(*
SPDX-FileCopyrightText: c 2026 Oleksandr Tiutyk <trofimich@gmail.com>
SPDX-License-Identifier: MIT
License: https://opensource.org/license/mit
*)

(*!
<summary>Checks that a long aggregate diagnostic is terminated and ends in an ellipsis.</summary>
<description>
Uses one task and stays at a stable address while assertions are bound to this instance.
</description>
*)

{attribute 'no_assign'}
{attribute 'no_explicit_call' := 'do not call this function block directly'}
FUNCTION_BLOCK AggregateExceptionBoundedMessageTest EXTENDS TOF_Testing.SingleCycleTest
VAR_STAT
	{attribute 'hide'}
	_ClassName : STRING := __POUNAME();
END_VAR
VAR
	_Aggregate : TOF_Core.AggregateException;
END_VAR

(*!
<summary>Checks that a long aggregate diagnostic is terminated and ends in an ellipsis.</summary>
<description>
Three entries share one task-managed cause. Each payload fills half the diagnostic buffer so the
combined message exceeds its capacity. The persistent reference array is released in AfterTest.
</description>
*)
METHOD PROTECTED ExecuteTest
VAR
	exceptionCode : __SYSTEM.ExceptionCode;
	caught : TOF_Core.IException;
	cause : TOF_Core.IStandardException;
	payload : TOF_Core.ERROR_MESSAGE;
	message : TOF_Core.ERROR_MESSAGE;
	payloadUnits : POINTER TO WORD;
	messageUnits : POINTER TO WORD;
	i : UDINT;
END_VAR
VAR CONSTANT
	MESSAGE_CAPACITY : UDINT := TOF_Core.Parameters.ERROR_MESSAGE_WIDE_CHAR_SIZE;
END_VAR
// Make an ASCII payload whose length scales with the documented diagnostic capacity.
payloadUnits := ADR(payload);

FOR i := 0 TO MESSAGE_CAPACITY / 2 - 1 DO
	payloadUnits[i] := WORD#16#0058; // Uppercase X makes the retained prefix distinguishable from the ellipsis.
END_FOR

payloadUnits[MESSAGE_CAPACITY / 2] := TO_WORD(TOF_Core.UnsignedInt16.MIN_VALUE);

// Obtain one dynamic cause so repeated entries exercise permitted sharing.
__TRY
	TOF_Core.Exceptions.ThrowStandard(
		sourceNamespaceName := NamespaceName,
		sourceClassName := ClassName,
		sourcePOUName := __POUNAME(),
		sourcePosition := __POSITION(),
		message := payload
	);
__CATCH(exceptionCode)
	caught := TOF_Core.ExceptionManager.GetLastException(
		exceptionCode := exceptionCode,
		catchPointNamespaceName := NamespaceName,
		catchPointPOUName := __POUNAME(),
		catchPointPosition := __POSITION()
	);
__ENDTRY

IF NOT __QUERYINTERFACE(caught, cause) THEN
	RecordFailure(message := "A task-owned payload is required for the aggregate length check");
	RETURN;
END_IF

_Aggregate.AddInnerException(innerException := cause);
_Aggregate.AddInnerException(innerException := cause);
_Aggregate.AddInnerException(innerException := cause);
message := _Aggregate.GetMessage();

messageUnits := ADR(message);

IF messageUnits[MESSAGE_CAPACITY] <> TO_WORD(TOF_Core.UnsignedInt16.MIN_VALUE) THEN
	RecordFailure(message := "The last storage unit must terminate the aggregate diagnostic");
	RETURN;
END_IF

Assert.ThatUDInt(
	actual := TOF_Core.WideStrings.GetLength(value := message),
	message := "The bounded aggregate message must fill the available character capacity"
).ToBe(expected := MESSAGE_CAPACITY);
Assert.ThatBool(
	actual := Tc2_Standard.WFIND(STR1 := message, STR2 := "3 aggregated exceptions$R0:") = 1,
	message := "The bounded message must retain the aggregate header and the first entry marker"
).IsTrue();
Assert.ThatBool(
	actual := messageUnits[MESSAGE_CAPACITY - 2] = WORD#16#0058,
	message := "The bounded message must retain cause text immediately before the ellipsis"
).IsTrue();
Assert.ThatBool(
	actual := messageUnits[MESSAGE_CAPACITY - 1] = TOF_Core.WideStrings.ELLIPSIS,
	message := "The final character must be an ellipsis"
).IsTrue();
END_METHOD

(*!
<summary>Clears the caller-owned aggregate storage before the result is reported.</summary>
<description>
Safe after partial setup or repeated Clear. The task memory manager retains ownership of dynamic causes.
</description>
*)
METHOD PROTECTED AfterTest
_Aggregate.Clear();
END_METHOD

//! <summary>Borrows the concrete class name. Callers must not modify it.</summary>
{attribute 'monitoring' := 'call'}
PROPERTY ClassName : REFERENCE TO STRING
GET
ClassName REF= _ClassName;
END_GET
END_PROPERTY

//! <summary>Borrows the compiler-initialized namespace name. Callers must not modify it.</summary>
{attribute 'monitoring' := 'call'}
PROPERTY NamespaceName : REFERENCE TO STRING
GET
NamespaceName REF= CurrentNamespace.Name;
END_GET
END_PROPERTY

//! <summary>Reports the concrete instance size in bytes.</summary>
{attribute 'monitoring' := 'call'}
PROPERTY SelfSize : ULINT
GET
SelfSize := XSIZEOF(THIS^);
END_GET
END_PROPERTY

END_FUNCTION_BLOCK

(* stored: Version 1.1.0.1
   POU AggregateExceptionBoundedMessageTest: Id {2554335a-8f4c-431b-bf31-5e17f62834b8}, SpecialFunc None
   Method ExecuteTest: Id {c925eba0-3c06-43e8-8fe2-e661cff1b46a}
   Method AfterTest: Id {da596345-5a78-4729-b445-ef794f46aef9}
   Property ClassName: Id {0583e574-cfb6-4c76-9ded-1b12e65bf318}
   Get Get: Id {60d99622-b8b3-4d56-bc98-16b9192d666d}
   Property NamespaceName: Id {55078304-e630-4323-b2a4-adce39836f0b}
   Get Get: Id {ffa225cd-9c4e-49be-a96b-9778e1e0b8e5}
   Property SelfSize: Id {decd74a7-f436-4301-9d3b-ac96926ad372}
   Get Get: Id {3cbe2884-d542-4cb8-b882-6634e08f5dda} *)
